// SIMATIC S7-200 project (STEP 7-Micro/WIN), CPU 224 CN REL 02.01

SYMBOL_TABLE 用户定义1
顶料到位检测           I0.0
顶料复位检测           I0.1
推料到位检测           I0.2
推料复位检测           I0.3
物料台物料检测          I0.4
物料不够检测           I0.5
物料有无检测           I0.6
金属传感器检测          I0.7
推料按钮             I1.2
启动按钮             I1.3
急停按钮             I1.4
单机全线             I1.5
准备就绪             M0.0
启动               M0.1
顶料电磁阀            Q0.0
推料电磁阀            Q0.1
正常工作指示           Q0.7
推料完成指示           Q1.0
红色指示灯            Q1.1
供料请求             V1000.4
网络正常             V1010.0
全线模式             V1010.1
料不足              V1010.2
缺料               V1010.3
供料完成             V1010.4
END_SYMBOL_TABLE

ORGANIZATION_BLOCK 主程序:OB1
TITLE=程序注释
BEGIN
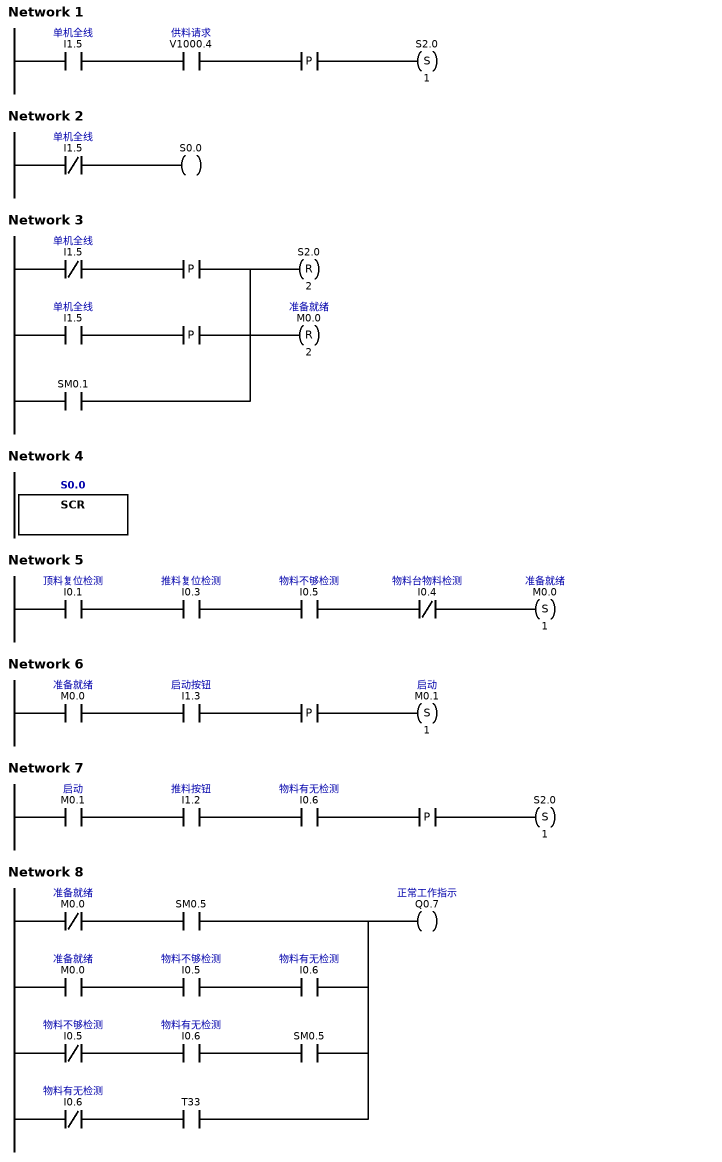
Network 1
LD     单机全线:I1.5
A      供料请求:V1000.4
EU
S      S2.0, 1
Network 2
LDN    单机全线:I1.5
=      S0.0
Network 3
LDN    单机全线:I1.5
EU
LD     单机全线:I1.5
EU
OLD
O      SM0.1
R      S2.0, 2
R      准备就绪:M0.0, 2
Network 4
LSCR   S0.0
Network 5
LD     顶料复位检测:I0.1
A      推料复位检测:I0.3
A      物料不够检测:I0.5
AN     物料台物料检测:I0.4
S      准备就绪:M0.0, 1
Network 6
LD     准备就绪:M0.0
A      启动按钮:I1.3
EU
S      启动:M0.1, 1
Network 7
LD     启动:M0.1
A      推料按钮:I1.2
A      物料有无检测:I0.6
EU
S      S2.0, 1
Network 8
LDN    准备就绪:M0.0
A      SM0.5
LD     准备就绪:M0.0
A      物料不够检测:I0.5
A      物料有无检测:I0.6
OLD
LDN    物料不够检测:I0.5
A      物料有无检测:I0.6
A      SM0.5
OLD
LDN    物料有无检测:I0.6
A      T33
OLD
=      正常工作指示:Q0.7
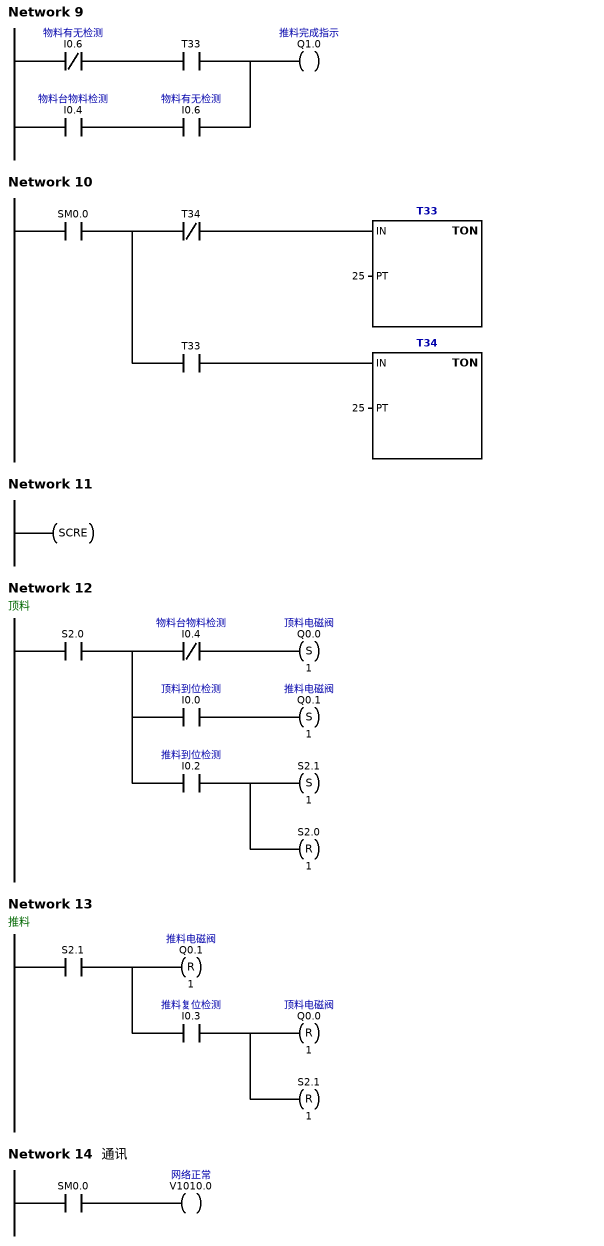
Network 9
LDN    物料有无检测:I0.6
A      T33
LD     物料台物料检测:I0.4
A      物料有无检测:I0.6
OLD
=      推料完成指示:Q1.0
Network 10
LD     SM0.0
LPS
AN     T34
TON    T33, 25
LPP
A      T33
TON    T34, 25
Network 11
SCRE
Network 12
// 顶料
LD     S2.0
LPS
AN     物料台物料检测:I0.4
S      顶料电磁阀:Q0.0, 1
LRD
A      顶料到位检测:I0.0
S      推料电磁阀:Q0.1, 1
LPP
A      推料到位检测:I0.2
S      S2.1, 1
R      S2.0, 1
Network 13
// 推料
LD     S2.1
R      推料电磁阀:Q0.1, 1
A      推料复位检测:I0.3
R      顶料电磁阀:Q0.0, 1
R      S2.1, 1
Network 14 // 通讯
LD     SM0.0
=      网络正常:V1010.0
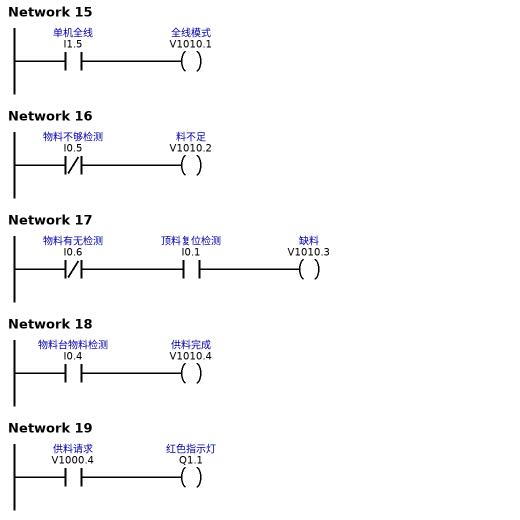
Network 15
LD     单机全线:I1.5
=      全线模式:V1010.1
Network 16
LDN    物料不够检测:I0.5
=      料不足:V1010.2
Network 17
LDN    物料有无检测:I0.6
A      顶料复位检测:I0.1
=      缺料:V1010.3
Network 18
LD     物料台物料检测:I0.4
=      供料完成:V1010.4
Network 19
LD     供料请求:V1000.4
=      红色指示灯:Q1.1
END_ORGANIZATION_BLOCK
